FUNCTION_BLOCK FB_Gr00ManualInit
(*

The function block used to initialize manual mode.

Constructor: 		Patryk Panylo
Company:		E. Riexinger GmbH
Date:			28.04.2015
Version:			1.00

Date:			Revision:		Who:				Comment
dd.mm.yyyy		x.xx			Initials			comment

*)
VAR_INPUT
	(* Input variables / Eingang Variablen *)
	bFirstTime					:BOOL;
END_VAR
VAR_OUTPUT
	(* Output variables / Ausgang Variablen *)

END_VAR
VAR_IN_OUT
	(* Input Output variables / Ausgang Variablen *)

END_VAR
VAR
	(* Enummerations *)

	(* Variables *)

	(* References *)

	(* Interfaces *)

	(* Instances *)

END_VAR


(* Initializing variables *)
IF NOT bFirstTime
THEN
	(* Program init *)
	Gr00Control.fbProgram.bRead := FALSE;								(* Read program *)

	(* Manual procedure *)
	Gr00Manual.fbProcedure.bEnable := FALSE;							(* Start init process *)
	Gr00Manual.fbProcedure.bExecute := FALSE;
	Gr00Manual.fbProcedure();

	bFirstTime := TRUE;
END_IF;

END_FUNCTION_BLOCK

(* stored: Version 1.1.0.1, ProductVersion 3.1.4024.15
   POU FB_Gr00ManualInit: Id {b947fd95-b559-41ef-87f8-b767781cbdb1}, SpecialFunc None *)
